FUNCTION_BLOCK FrequenciaSel (* Frequencia do motor: do ATV (REAL, Hz) ou da Sulzer (INT, 0,1 Hz) *)
  (* Standard: 61499-2 *)
  (* Version 1.0, 04/11/2026, Hidryco, Hidryco, 1.0: REQ_REAL repassa FreqReal; REQ_HZ10 converte FreqHz10 / 10. Vale o ultimo que chegou (cada motor so tem uma das duas ligadas no hardware). *)
  PACKAGE SE.Nereda;
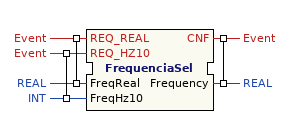
  EVENT_INPUT
    REQ_REAL WITH FreqReal; (* Frequencia em Hz (symlink MotorFrequecy) *)
    REQ_HZ10 WITH FreqHz10; (* Frequencia em 0,1 Hz (symlink FreqHz10, Sulzer) *)
  END_EVENT
  EVENT_OUTPUT
    CNF WITH Frequency; (* Frequencia em Hz *)
  END_EVENT
  VAR_INPUT
    FreqReal : REAL; (* Hz *)
    FreqHz10 : INT; (* 0,1 Hz *)
  END_VAR
  VAR_OUTPUT
    Frequency : REAL; (* Hz *)
  END_VAR
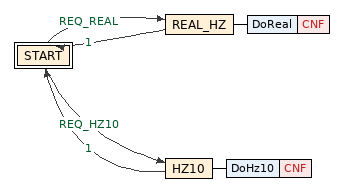
  EC_STATES
    START; (* Estado inicial *)
    REAL_HZ : DoReal -> CNF; (* Do ATV *)
    HZ10 : DoHz10 -> CNF; (* Da Sulzer *)
  END_STATES
  EC_TRANSITIONS
    START TO REAL_HZ := REQ_REAL;
    REAL_HZ TO START := 1;
    START TO HZ10 := REQ_HZ10;
    HZ10 TO START := 1;
  END_TRANSITIONS
  ALGORITHM DoReal IN ST: (* Hz direto *)
Frequency := FreqReal;
  END_ALGORITHM
  ALGORITHM DoHz10 IN ST: (* 0,1 Hz para Hz *)
Frequency := INT_TO_REAL(FreqHz10) / 10.0;
  END_ALGORITHM
END_FUNCTION_BLOCK
